TYPE ST_CommonConfig_REAL :
STRUCT
	value	: REAL;
	is_available : UDINT;
END_STRUCT
END_TYPE

(* stored: Version 1.1.0.1, ProductVersion 3.1.4024.12
   DUT ST_CommonConfig_REAL: Id {b1921432-4ca8-4785-ad34-281873a13505} *)
